Fanuc KAREL source: KX00028.KL

PROGRAM KX00028
%NOLOCKGROUP
%TIMESLICE = 8
VAR
  I: INTEGER
  J: INTEGER
  B: BOOLEAN
  F: FILE
  S: STRING[80]
  P: XYZWPR
BEGIN
  I = 1
END KX00028
